FUNCTION_BLOCK FB_CIP_ClientTank EXTENDS FB_SFC_Cycle IMPLEMENTS ITF_FB_SFC_Cycle
VAR_INPUT	
	valTank_A				: E_Pis_Name;
	valTank_A_Sprinkler		: E_Pis_Name;
	valTank_A_Main			: E_Pis_Name;
	valTank_B				: E_Pis_Name;
	valTank_B_Sprinkler		: E_Pis_Name;	
	valTank_B_Main			: E_Pis_Name;	
	valDrain				: E_Pis_Name;
END_VAR
VAR_OUTPUT
END_VAR
VAR

	eReq				: E_CIP_ClientTank;
	eProcess			: E_CIP_ClientTank;
	eStatus				: E_CIP_ClientTank;
	
	fbPis					: FB_Piston;
	stPis_Tank_A			: REFERENCE TO ST_Piston;
	stPis_Tank_A_Sprinkler	: REFERENCE TO ST_Piston;
	stPis_Tank_A_Main		: REFERENCE TO ST_Piston;
	stPis_Tank_B			: REFERENCE TO ST_Piston;
	stPis_Tank_B_Sprinkler	: REFERENCE TO ST_Piston;
	stPis_Tank_B_Main		: REFERENCE TO ST_Piston;
	stPis_Drain				: REFERENCE TO ST_Piston;

	tonDrainTime: TON;
	rt_Req_Reset: R_TRIG;
END_VAR
VAR_IN_OUT


END_VAR

act_GetReference();

act_Oper();
IF NOT Init.x THEN;
	act_Status();
END_IF

tonDrainTime(PT:=T#1M, IN:=eStatus=E_CIP_ClientTank.eDrain);
IF tonDrainTime.Q 
AND eReq=E_CIP_ClientTank.eNone
AND eProcess=E_CIP_ClientTank.eNone
THEN;
	eReq:=E_CIP_ClientTank.eClose;
END_IF

m_Request_Reset(memo:=rt_Req_Reset);

ACTION _aClose_active:
bStepDone:=FALSE;
IF TRUE 
AND eStatus=E_CIP_ClientTank.eClose
THEN;
	bStepDone:=TRUE;
END_IF
END_ACTION

ACTION _aClose_entry:
fbPis.m_SetByRecipe(stPis:=stPis_Tank_A, 				req:=E_Piston_Recipe_State.Release);
fbPis.m_SetByRecipe(stPis:=stPis_Tank_A_Sprinkler, 		req:=E_Piston_Recipe_State.Release);
fbPis.m_SetByRecipe(stPis:=stPis_Tank_A_Main, 			req:=E_Piston_Recipe_State.Release);
fbPis.m_SetByRecipe(stPis:=stPis_Tank_B, 				req:=E_Piston_Recipe_State.Release);
fbPis.m_SetByRecipe(stPis:=stPis_Tank_B_Sprinkler, 		req:=E_Piston_Recipe_State.Release);
fbPis.m_SetByRecipe(stPis:=stPis_Tank_B_Main, 			req:=E_Piston_Recipe_State.Release);
fbPis.m_SetByRecipe(stPis:=stPis_Drain, 				req:=E_Piston_Recipe_State.Release);
END_ACTION

ACTION _aDone_entry:
eProcess:=E_CIP_ClientTank.eNone;
eReq:=E_CIP_ClientTank.eNone;
bRun:=FALSE;
bDone:=TRUE;
END_ACTION

ACTION _aDrain_active:
bStepDone:=FALSE;
IF TRUE 
AND eStatus=E_CIP_ClientTank.eDrain
THEN;
	bStepDone:=TRUE;
END_IF
END_ACTION

ACTION _aDrain_entry:
fbPis.m_SetByRecipe(stPis:=stPis_Tank_A, 				req:=E_Piston_Recipe_State.Release);
fbPis.m_SetByRecipe(stPis:=stPis_Tank_A_Sprinkler, 		req:=E_Piston_Recipe_State.Release);
fbPis.m_SetByRecipe(stPis:=stPis_Tank_A_Main, 			req:=E_Piston_Recipe_State.Release);
fbPis.m_SetByRecipe(stPis:=stPis_Tank_B, 				req:=E_Piston_Recipe_State.Release);
fbPis.m_SetByRecipe(stPis:=stPis_Tank_B_Sprinkler, 		req:=E_Piston_Recipe_State.Release);
fbPis.m_SetByRecipe(stPis:=stPis_Tank_B_Main, 			req:=E_Piston_Recipe_State.Release);
fbPis.m_SetByRecipe(stPis:=stPis_Drain, 				req:=E_Piston_Recipe_State.Act);
END_ACTION

ACTION _aInit_active:
SFCReset:=FALSE;
END_ACTION

ACTION _aInit_exit:
eProcess:=E_CIP_ClientTank.eNone;
eReq:=E_CIP_ClientTank.eNone;
END_ACTION

ACTION _aReady_active:


CASE eReq OF
	E_CIP_ClientTank.eClose:;
			IF TRUE THEN;
				eProcess:=E_CIP_ClientTank.eClose;
			END_IF

	E_CIP_ClientTank.eTank_A:;
			IF TRUE THEN;
				eProcess:=E_CIP_ClientTank.eTank_A;
			END_IF	
			
	E_CIP_ClientTank.eTank_A_Sprinkler:;
			IF TRUE THEN;
				eProcess:=E_CIP_ClientTank.eTank_A_Sprinkler;
			END_IF
			
	E_CIP_ClientTank.eTank_B:;
			IF TRUE THEN;
				eProcess:=E_CIP_ClientTank.eTank_B;
			END_IF	
	
	E_CIP_ClientTank.eTank_B_Sprinkler:;
			IF TRUE THEN;
				eProcess:=E_CIP_ClientTank.eTank_B_Sprinkler;
			END_IF	

	E_CIP_ClientTank.eDrain:;
			IF TRUE THEN;
				eProcess:=E_CIP_ClientTank.eDrain;
			END_IF	
	

END_CASE
END_ACTION

ACTION _aReady_exit:
bRun:=TRUE;
bDone:=FALSE;
END_ACTION

ACTION _aTank_A_active:
bStepDone:=FALSE;
IF TRUE 
AND eStatus=E_CIP_ClientTank.eTank_A
THEN;
	bStepDone:=TRUE;
END_IF
END_ACTION

ACTION _aTank_A_entry:
fbPis.m_SetByRecipe(stPis:=stPis_Tank_A, 				req:=E_Piston_Recipe_State.Act);
fbPis.m_SetByRecipe(stPis:=stPis_Tank_A_Sprinkler, 		req:=E_Piston_Recipe_State.Release);
fbPis.m_SetByRecipe(stPis:=stPis_Tank_A_Main, 			req:=E_Piston_Recipe_State.Release);
fbPis.m_SetByRecipe(stPis:=stPis_Tank_B, 				req:=E_Piston_Recipe_State.Release);
fbPis.m_SetByRecipe(stPis:=stPis_Tank_B_Sprinkler, 		req:=E_Piston_Recipe_State.Release);
fbPis.m_SetByRecipe(stPis:=stPis_Tank_B_Main, 			req:=E_Piston_Recipe_State.Release);
fbPis.m_SetByRecipe(stPis:=stPis_Drain, 				req:=E_Piston_Recipe_State.Release);
END_ACTION

ACTION _aTank_A_Sprinkler_active:
bStepDone:=FALSE;
IF TRUE 
AND eStatus=E_CIP_ClientTank.eTank_A_Sprinkler
THEN;
	bStepDone:=TRUE;
END_IF
END_ACTION

ACTION _aTank_A_Sprinkler_entry:
fbPis.m_SetByRecipe(stPis:=stPis_Tank_A, 				req:=E_Piston_Recipe_State.Act);
fbPis.m_SetByRecipe(stPis:=stPis_Tank_A_Sprinkler, 		req:=E_Piston_Recipe_State.Act);
fbPis.m_SetByRecipe(stPis:=stPis_Tank_A_Main, 			req:=E_Piston_Recipe_State.Act);
fbPis.m_SetByRecipe(stPis:=stPis_Tank_B, 				req:=E_Piston_Recipe_State.Release);
fbPis.m_SetByRecipe(stPis:=stPis_Tank_B_Sprinkler, 		req:=E_Piston_Recipe_State.Release);
fbPis.m_SetByRecipe(stPis:=stPis_Tank_B_Main, 			req:=E_Piston_Recipe_State.Release);
fbPis.m_SetByRecipe(stPis:=stPis_Drain, 				req:=E_Piston_Recipe_State.Release);
END_ACTION

ACTION _aTank_B_active:
bStepDone:=FALSE;
IF TRUE 
AND eStatus=E_CIP_ClientTank.eTank_B
THEN;
	bStepDone:=TRUE;
END_IF
END_ACTION

ACTION _aTank_B_entry:
fbPis.m_SetByRecipe(stPis:=stPis_Tank_A, 				req:=E_Piston_Recipe_State.Release);
fbPis.m_SetByRecipe(stPis:=stPis_Tank_A_Sprinkler, 		req:=E_Piston_Recipe_State.Release);
fbPis.m_SetByRecipe(stPis:=stPis_Tank_A_Main, 			req:=E_Piston_Recipe_State.Release);
fbPis.m_SetByRecipe(stPis:=stPis_Tank_B, 				req:=E_Piston_Recipe_State.Act);
fbPis.m_SetByRecipe(stPis:=stPis_Tank_B_Sprinkler, 		req:=E_Piston_Recipe_State.Release);
fbPis.m_SetByRecipe(stPis:=stPis_Tank_B_Main, 			req:=E_Piston_Recipe_State.Release);
fbPis.m_SetByRecipe(stPis:=stPis_Drain, 				req:=E_Piston_Recipe_State.Release);
END_ACTION

ACTION _aTank_B_Sprinkler_active:
bStepDone:=FALSE;
IF TRUE 
AND eStatus=E_CIP_ClientTank.eTank_B_Sprinkler
THEN;
	bStepDone:=TRUE;
END_IF
END_ACTION

ACTION _aTank_B_Sprinkler_entry:
fbPis.m_SetByRecipe(stPis:=stPis_Tank_A, 				req:=E_Piston_Recipe_State.Release);
fbPis.m_SetByRecipe(stPis:=stPis_Tank_A_Sprinkler, 		req:=E_Piston_Recipe_State.Release);
fbPis.m_SetByRecipe(stPis:=stPis_Tank_A_Main, 			req:=E_Piston_Recipe_State.Release);
fbPis.m_SetByRecipe(stPis:=stPis_Tank_B, 				req:=E_Piston_Recipe_State.Act);
fbPis.m_SetByRecipe(stPis:=stPis_Tank_B_Sprinkler, 		req:=E_Piston_Recipe_State.Act);
fbPis.m_SetByRecipe(stPis:=stPis_Tank_B_Main, 			req:=E_Piston_Recipe_State.Act);
fbPis.m_SetByRecipe(stPis:=stPis_Drain, 				req:=E_Piston_Recipe_State.Release);
END_ACTION

ACTION act_GetReference:
m_Set_SFCFlags_Reference();
	
stPis_Tank_A				REF= g_Piston.stPis[valTank_A];
stPis_Tank_A_Sprinkler		REF= g_Piston.stPis[valTank_A_Sprinkler];
stPis_Tank_A_Main			REF= g_Piston.stPis[valTank_A_Main];
stPis_Tank_B				REF= g_Piston.stPis[valTank_B];
stPis_Tank_B_Sprinkler		REF= g_Piston.stPis[valTank_B_Sprinkler];
stPis_Tank_B_Main			REF= g_Piston.stPis[valTank_B_Main];
stPis_Drain					REF= g_Piston.stPis[valDrain];
END_ACTION

ACTION act_Oper:
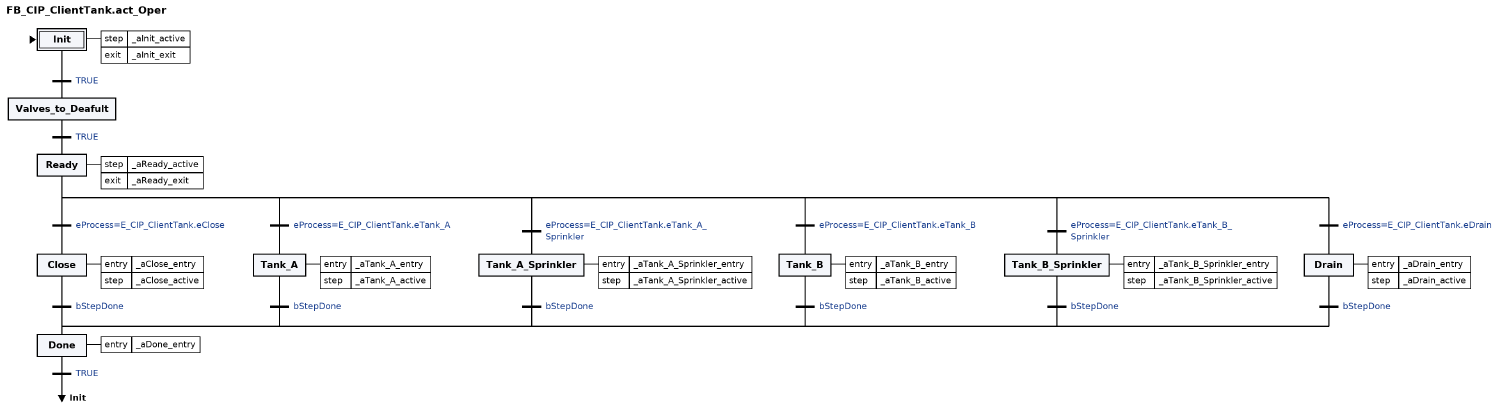
INITIAL_STEP Init:  // min time T#0.5s
    _aInit_active(N);  // step action
    _aInit_exit(P0);  // exit action
END_STEP
TRANSITION FROM Init TO Valves_to_Deafult
    := TRUE;
END_TRANSITION
STEP Valves_to_Deafult:
END_STEP
TRANSITION FROM Valves_to_Deafult TO Ready
    := TRUE;
END_TRANSITION
STEP Ready:
    _aReady_active(N);  // step action
    _aReady_exit(P0);  // exit action
END_STEP
TRANSITION FROM Ready TO Close
    := eProcess=E_CIP_ClientTank.eClose;
END_TRANSITION
STEP Close:
    _aClose_entry(P1);  // entry action
    _aClose_active(N);  // step action
END_STEP
TRANSITION FROM Close TO Done
    := bStepDone;
END_TRANSITION
TRANSITION FROM Ready TO Tank_A
    := eProcess=E_CIP_ClientTank.eTank_A;
END_TRANSITION
STEP Tank_A:
    _aTank_A_entry(P1);  // entry action
    _aTank_A_active(N);  // step action
END_STEP
TRANSITION FROM Tank_A TO Done
    := bStepDone;
END_TRANSITION
TRANSITION FROM Ready TO Tank_A_Sprinkler
    := eProcess=E_CIP_ClientTank.eTank_A_Sprinkler;
END_TRANSITION
STEP Tank_A_Sprinkler:
    _aTank_A_Sprinkler_entry(P1);  // entry action
    _aTank_A_Sprinkler_active(N);  // step action
END_STEP
TRANSITION FROM Tank_A_Sprinkler TO Done
    := bStepDone;
END_TRANSITION
TRANSITION FROM Ready TO Tank_B
    := eProcess=E_CIP_ClientTank.eTank_B;
END_TRANSITION
STEP Tank_B:
    _aTank_B_entry(P1);  // entry action
    _aTank_B_active(N);  // step action
END_STEP
TRANSITION FROM Tank_B TO Done
    := bStepDone;
END_TRANSITION
TRANSITION FROM Ready TO Tank_B_Sprinkler
    := eProcess=E_CIP_ClientTank.eTank_B_Sprinkler;
END_TRANSITION
STEP Tank_B_Sprinkler:
    _aTank_B_Sprinkler_entry(P1);  // entry action
    _aTank_B_Sprinkler_active(N);  // step action
END_STEP
TRANSITION FROM Tank_B_Sprinkler TO Done
    := bStepDone;
END_TRANSITION
TRANSITION FROM Ready TO Drain
    := eProcess=E_CIP_ClientTank.eDrain;
END_TRANSITION
STEP Drain:
    _aDrain_entry(P1);  // entry action
    _aDrain_active(N);  // step action
END_STEP
TRANSITION FROM Drain TO Done
    := bStepDone;
END_TRANSITION
STEP Done:  // min time T#0.2s
    _aDone_entry(P1);  // entry action
END_STEP
TRANSITION FROM Done TO Init
    := TRUE;
END_TRANSITION
// branch label Branch2_act_Oper
END_ACTION

ACTION act_Status:
IF bReady AND bDone OR TRUE THEN;
	IF TRUE 
	AND fbPis.m_CheckByRecipe(stPis:=stPis_Tank_A, 				req:=E_Piston_Recipe_State.Release)
	AND fbPis.m_CheckByRecipe(stPis:=stPis_Tank_A_Sprinkler, 	req:=E_Piston_Recipe_State.Release)
	AND fbPis.m_CheckByRecipe(stPis:=stPis_Tank_A_Main, 		req:=E_Piston_Recipe_State.Release)
	AND fbPis.m_CheckByRecipe(stPis:=stPis_Tank_B, 				req:=E_Piston_Recipe_State.Release)
	AND fbPis.m_CheckByRecipe(stPis:=stPis_Tank_B_Sprinkler, 	req:=E_Piston_Recipe_State.Release)
	AND fbPis.m_CheckByRecipe(stPis:=stPis_Tank_B_Main, 		req:=E_Piston_Recipe_State.Release)
	AND fbPis.m_CheckByRecipe(stPis:=stPis_Drain, 				req:=E_Piston_Recipe_State.Release)
	THEN;
		eStatus:=E_CIP_ClientTank.eClose;
		
	ELSIF TRUE 
	AND fbPis.m_CheckByRecipe(stPis:=stPis_Tank_A, 				req:=E_Piston_Recipe_State.Act)
	AND fbPis.m_CheckByRecipe(stPis:=stPis_Tank_A_Sprinkler, 	req:=E_Piston_Recipe_State.Release)
	AND fbPis.m_CheckByRecipe(stPis:=stPis_Tank_A_Main, 		req:=E_Piston_Recipe_State.Release)
	AND fbPis.m_CheckByRecipe(stPis:=stPis_Tank_B, 				req:=E_Piston_Recipe_State.Release)
	AND fbPis.m_CheckByRecipe(stPis:=stPis_Tank_B_Sprinkler, 	req:=E_Piston_Recipe_State.Release)
	AND fbPis.m_CheckByRecipe(stPis:=stPis_Tank_B_Main, 		req:=E_Piston_Recipe_State.Release)
	AND fbPis.m_CheckByRecipe(stPis:=stPis_Drain, 				req:=E_Piston_Recipe_State.Release)
	THEN;
		eStatus:=E_CIP_ClientTank.eTank_A;
	
	ELSIF TRUE 
	AND fbPis.m_CheckByRecipe(stPis:=stPis_Tank_A, 				req:=E_Piston_Recipe_State.Act)
	AND fbPis.m_CheckByRecipe(stPis:=stPis_Tank_A_Sprinkler, 	req:=E_Piston_Recipe_State.Act)
	AND fbPis.m_CheckByRecipe(stPis:=stPis_Tank_A_Main, 		req:=E_Piston_Recipe_State.Act)
	AND fbPis.m_CheckByRecipe(stPis:=stPis_Tank_B, 				req:=E_Piston_Recipe_State.Release)
	AND fbPis.m_CheckByRecipe(stPis:=stPis_Tank_B_Sprinkler, 	req:=E_Piston_Recipe_State.Release)
	AND fbPis.m_CheckByRecipe(stPis:=stPis_Tank_B_Main, 		req:=E_Piston_Recipe_State.Release)
	AND fbPis.m_CheckByRecipe(stPis:=stPis_Drain, 				req:=E_Piston_Recipe_State.Release)
	THEN;
		eStatus:=E_CIP_ClientTank.eTank_A_Sprinkler;
		
	ELSIF TRUE 
	AND fbPis.m_CheckByRecipe(stPis:=stPis_Tank_A, 				req:=E_Piston_Recipe_State.Release)
	AND fbPis.m_CheckByRecipe(stPis:=stPis_Tank_A_Sprinkler, 	req:=E_Piston_Recipe_State.Release)
	AND fbPis.m_CheckByRecipe(stPis:=stPis_Tank_A_Main, 		req:=E_Piston_Recipe_State.Release)
	AND fbPis.m_CheckByRecipe(stPis:=stPis_Tank_B, 				req:=E_Piston_Recipe_State.Act)
	AND fbPis.m_CheckByRecipe(stPis:=stPis_Tank_B_Sprinkler, 	req:=E_Piston_Recipe_State.Release)
	AND fbPis.m_CheckByRecipe(stPis:=stPis_Tank_B_Main, 		req:=E_Piston_Recipe_State.Release)
	AND fbPis.m_CheckByRecipe(stPis:=stPis_Drain, 				req:=E_Piston_Recipe_State.Release)
	THEN;
		eStatus:=E_CIP_ClientTank.eTank_B;	
		
	ELSIF TRUE 
	AND fbPis.m_CheckByRecipe(stPis:=stPis_Tank_A, 				req:=E_Piston_Recipe_State.Release)
	AND fbPis.m_CheckByRecipe(stPis:=stPis_Tank_A_Sprinkler, 	req:=E_Piston_Recipe_State.Release)
	AND fbPis.m_CheckByRecipe(stPis:=stPis_Tank_A_Main, 		req:=E_Piston_Recipe_State.Release)
	AND fbPis.m_CheckByRecipe(stPis:=stPis_Tank_B, 				req:=E_Piston_Recipe_State.Act)
	AND fbPis.m_CheckByRecipe(stPis:=stPis_Tank_B_Sprinkler, 	req:=E_Piston_Recipe_State.Act)
	AND fbPis.m_CheckByRecipe(stPis:=stPis_Tank_B_Main, 		req:=E_Piston_Recipe_State.Act)
	AND fbPis.m_CheckByRecipe(stPis:=stPis_Drain, 				req:=E_Piston_Recipe_State.Release)
	THEN;
		eStatus:=E_CIP_ClientTank.eTank_B_Sprinkler;
		
	ELSIF TRUE 	
	AND fbPis.m_CheckByRecipe(stPis:=stPis_Tank_A, 				req:=E_Piston_Recipe_State.Release)
	AND fbPis.m_CheckByRecipe(stPis:=stPis_Tank_A_Sprinkler, 	req:=E_Piston_Recipe_State.Release)
	AND fbPis.m_CheckByRecipe(stPis:=stPis_Tank_A_Main, 		req:=E_Piston_Recipe_State.Release)
	AND fbPis.m_CheckByRecipe(stPis:=stPis_Tank_B, 				req:=E_Piston_Recipe_State.Release)
	AND fbPis.m_CheckByRecipe(stPis:=stPis_Tank_B_Sprinkler, 	req:=E_Piston_Recipe_State.Release)
	AND fbPis.m_CheckByRecipe(stPis:=stPis_Tank_B_Main, 		req:=E_Piston_Recipe_State.Release)
	AND fbPis.m_CheckByRecipe(stPis:=stPis_Drain, 				req:=E_Piston_Recipe_State.Act)
	THEN;
		eStatus:=E_CIP_ClientTank.eDrain;
		
	ELSE;
		eStatus:=E_CIP_ClientTank.eNone;
	END_IF
ELSE;
	eStatus:=E_CIP_ClientTank.eNone;
END_IF
END_ACTION

METHOD m_CheckStatus : BOOL
VAR_INPUT
	eReqStatus		: E_CIP_ClientTank;
END_VAR
IF eStatus=eReqStatus 
AND eProcess=E_CIP_ClientTank.eNone
AND eReq=E_CIP_ClientTank.eNone
AND bReady
AND bDone
AND NOT bRun
THEN;
	m_CheckStatus:=TRUE;
END_IF
END_METHOD

METHOD m_Request_Reset : BOOL
VAR_IN_OUT
	memo: R_TRIG;
END_VAR
memo(CLK:=eReq=0);
IF TRUE 
AND memo.Q
THEN;
	SFCReset:=TRUE;
END_IF
END_METHOD

METHOD m_Run : BOOL
VAR_INPUT
	eReqProc			: E_CIP_ClientTank;
END_VAR
IF eProcess=E_CIP_ClientTank.eNone THEN;
	eProcess:=eReq:=eReqProc;
	bDone:=FALSE;
	m_Run:=TRUE;
END_IF
END_METHOD

METHOD m_Set_SFCFlags_Reference : BOOL
//Set reference to SFC flags

refSFC.SFCInit REF= SFCInit;
refSFC.SFCReset REF= SFCReset;
refSFC.SFCError REF= SFCError;
refSFC.SFCEnableLimit REF= SFCEnableLimit;
refSFC.SFCErrorStep REF= SFCErrorStep;
refSFC.SFCErrorPOU REF= SFCErrorPOU;
refSFC.SFCQuitError REF= SFCQuitError;
refSFC.SFCPause REF= SFCPause;
refSFC.SFCTrans REF= SFCTrans;
refSFC.SFCCurrentStep REF= SFCCurrentStep;
refSFC.SFCTip REF= SFCTip;
refSFC.SFCTipMode REF= SFCTipMode;

// Cycle handle for SFC
m_SFC_Handle();
END_METHOD

END_FUNCTION_BLOCK

(* stored: Version 1.1.0.1, ProductVersion 3.1.4024.13
   POU FB_CIP_ClientTank: Id {ec4051e0-f8dc-45bc-bf46-7adcfec692af}, SpecialFunc None
   Folder Manage: Id {75407563-912d-4908-b651-2f1b671d8753}
   Action _aClose_active: Id {92f6b6d1-b589-4a20-bcda-89bf8146bb5b}
   Action _aClose_entry: Id {e7dae316-3ace-4522-92c2-0cffa79ad812}
   Action _aDone_entry: Id {7884b3c0-ec72-4080-ae05-f0a6b28907f3}
   Action _aDrain_active: Id {f6cebb11-b4ad-49db-9d93-c21a8948919a}
   Action _aDrain_entry: Id {9d6fa881-c60b-4a07-bb86-a9b166160530}
   Action _aInit_active: Id {07963cc4-97a0-40c4-8d4a-8860062e87ff}
   Action _aInit_exit: Id {855f3e65-7ea9-4b16-90c8-ef323d24f02d}
   Action _aReady_active: Id {b8a80171-ccbc-439a-bcf2-0bdb246c8206}
   Action _aReady_exit: Id {4a24de33-5094-4e27-95ae-6434e8ee7ad6}
   Action _aTank_A_active: Id {86ddce0d-560e-43e6-8013-13a99078bfa4}
   Action _aTank_A_entry: Id {951a57df-a15c-4fee-b116-bcded9db2564}
   Action _aTank_A_Sprinkler_active: Id {2c65f399-d21d-479b-899d-841f0928a544}
   Action _aTank_A_Sprinkler_entry: Id {ed5047a0-51f6-49a8-939a-5f79d7c9f6ce}
   Action _aTank_B_active: Id {6b4bc092-8ce6-4648-a8ff-ad164d214ca2}
   Action _aTank_B_entry: Id {117ef39d-0a17-4a6d-aa08-2189f1a3d8a8}
   Action _aTank_B_Sprinkler_active: Id {56c82813-2539-44fc-8a4c-1ad71d2afce5}
   Action _aTank_B_Sprinkler_entry: Id {1df2f61b-c379-4645-855b-7a9b92b02674}
   Action act_GetReference: Id {62ed5244-769e-4b64-a5c5-5f290efa2568}
   Action act_Oper: Id {d68978ed-0f1f-4eaa-bed5-19d4ace73904}
   Action act_Status: Id {ea2c6eb6-6b5f-44a7-aec7-310eecd35922}
   Method m_CheckStatus: Id {cd38da1d-87fa-4c25-8cd1-074243f17cb1}
   Method m_Request_Reset: Id {ea357b7e-42a7-4b81-9b8a-30befe36872d}
   Method m_Run: Id {ec4b68e6-5819-4865-ba29-867baa0dec5e}
   Method m_Set_SFCFlags_Reference: Id {7e38792a-dc64-4fa1-bbd1-b9c8a5df9f5d} *)
